(* IEC 61131-3 sources: sis-interlock-demo/src/POUs/Sis/F_SisLowMask, 2 files *)

(* ---- F_SisLowMask.decl.st ---- *)
// Назначение: маска младших битов 0..uiCount − 1: 0 — 0, 16 и больше — 16#FFFF.
// Автор:      kr0nsch
// Версия:     0.1.0
// Документ:   docs/DESIGN.md, раздел «8.2 Функции работы с битами»
// ВНИМАНИЕ:   код демонстрационный и не предназначен для систем безопасности. Реальная ПАЗ
//             требует определения SIL, сертифицированных аппаратных и программных средств
//             и валидации по ГОСТ Р МЭК 61511.
FUNCTION F_SisLowMask : WORD
VAR_INPUT
    uiCount : UINT;  // число младших битов
END_VAR

(* ---- F_SisLowMask.impl.st ---- *)
IF uiCount = 0 THEN
    F_SisLowMask := 0;
ELSIF uiCount >= GVL_Const.WORD_BITS THEN
    // сдвиг на разрядность и больше не определён — значение задаётся явно
    F_SisLowMask := GVL_Const.WORD_ALL;
ELSE
    // старшие биты 16#FFFF после сдвига влево — единицы; XOR оставляет младшие uiCount единиц
    F_SisLowMask := SHL(GVL_Const.WORD_ALL, uiCount) XOR GVL_Const.WORD_ALL;
END_IF
